Fanuc KAREL source: KT00493.KL

PROGRAM KT00493
%NOLOCKGROUP
VAR
  P1: XYZWPR
  P2: POSITION
  OUT: BOOLEAN
BEGIN
  P1.X = 1.0
  OUT = P1 >=< P2
END KT00493
